(* IEC 61131-3 sources: llm-plc-st-eval/data/processed_definitivo/gpt-4o-2024-08-06/C3/few_shot, 3 files *)

(* ---- ejec_1.st ---- *)
PROGRAM PRG_Conversion
VAR_INPUT
    btnMarcha : BOOL; (* Contacto NA en paralelo *)
    btnParo : BOOL; (* Contacto NC en serie *)
END_VAR
VAR_OUTPUT
    motor : BOOL; (* Bobina motor *)
    lampara : BOOL; (* Bobina lámpara *)
END_VAR
VAR
    T1 : TON; (* Temporizador TON *)
END_VAR

(* Serie = AND, paralelo = OR, contacto NC = NOT *)
motor := ((btnMarcha OR motor) AND NOT btnParo);

(* Temporizador TON activado por el motor *)
T1(IN := motor, PT := T#10S);

(* La lámpara se activa cuando el temporizador alcanza el tiempo preestablecido *)
lampara := T1.Q;
END_PROGRAM

(* ---- ejec_2.st ---- *)
PROGRAM PRG_Conversion
VAR
    btnMarcha : BOOL; (* Contacto NA en paralelo *)
    btnParo : BOOL; (* Contacto NC en serie *)
    motor : BOOL; (* Bobina motor *)
    lampara : BOOL; (* Bobina lámpara *)
    T1 : TON; (* Temporizador TON *)
END_VAR

(* Serie = AND, paralelo = OR, contacto NC = NOT *)
motor := ((btnMarcha OR motor) AND NOT btnParo);

(* Configuración y ejecución del temporizador TON *)
T1(IN := motor, PT := T#10S);

(* Activación de la lámpara cuando T1.Q es TRUE *)
lampara := T1.Q;
END_PROGRAM

(* ---- ejec_3.st ---- *)
PROGRAM PRG_Conversion
VAR
    btnMarcha : BOOL; (* Contacto NA en paralelo *)
    btnParo : BOOL; (* Contacto NC en serie *)
    motor : BOOL; (* Bobina motor *)
    lampara : BOOL; (* Bobina lámpara *)
    T1 : TON; (* Temporizador TON *)
END_VAR

(* Serie = AND, paralelo = OR, contacto NC = NOT *)
motor := ((btnMarcha OR motor) AND NOT btnParo);

(* Configuración del temporizador TON *)
T1(IN := motor, PT := T#10S);

(* La lámpara se enciende cuando el temporizador alcanza el tiempo preestablecido *)
lampara := T1.Q;
END_PROGRAM
